// TIA Portal V21 export
// export: Created 2026-10-12T11:32:16.9402514Z, ExportSetting WithDefaults, DisplayName Totally Integrated Automation Portal, DisplayVersion V21, DisplayName STEP 7 Professional, DisplayVersion V21, DisplayName STEP 7 Safety, DisplayVersion V21, DisplayName Tech WebApplication, DisplayVersion V21, DisplayName WinCC Basic/Comfort/Advanced, DisplayVersion V21, DisplayName WinCC Unified, DisplayVersion V21
DATA_BLOCK "DB_TCP_IP"   // DB12
{ S7_Optimized_Access := 'TRUE' }
VERSION : 0.1
// stored: AutoNumber true, DBAccessibleFromOPCUA true, IsOnlyStoredInLoadMemory false, IsRetainMemResEnabled false, IsWriteProtectedInAS false, MemoryReserve 100
   VAR
      "MY CONNECT DATA" { S7_SetPoint := 'True'} : TCON_IP_v4;
      "NO OF DONE" { S7_SetPoint := 'True'} : UDInt;
      "NO OF ERROR" : UDInt;
      "ERROR STATUS" : UDInt;
   END_VAR
BEGIN
END_DATA_BLOCK
